Staubli VAL3: setActive.pgx

program setActive(num x_nIndex)
begin
  safeTemp:sSPoint[x_nIndex].bActive=(bActive==true)
end
